FUNCTION_BLOCK FB_Gr01AutoAlarm
(*

The function block used to control alarms in manual mode.

Constructor: 		Patryk Panylo
Company:		E. Riexinger GmbH
Date:			28.04.2015
Version:			1.00

Date:			Revision:		Who:				Comment
dd.mm.yyyy		x.xx			Initials			comment

*)
VAR_INPUT
	(* Input variables / Eingang Variablen *)
	etMachineMode				:ET_MachineMode;			(* Machine mode *)
	etMachineState				:ET_MachineState;			(* Machine state *)
	bNoEStop					:BOOL;						(* Emergency stop *)
	bConfirmAlarm				:BOOL;						(* Confirm alarm *)
	dtDateTime 					:DATE_AND_TIME;			(* Actual date and time *)
	nFatalErrorMaxIdx				:INT;						(* Maximal index of  using alarms *)
	nErrorMaxIdx					:INT;						(* Maximal index of  using alarms *)
	nWarningMaxIdx				:INT;						(* Maximal index of  using alarms *)
	nMessageMaxIdx				:INT;						(* Maximal index of  using alarms *)
	nHintMaxIdx					:INT;						(* Maximal index of  using alarms *)
	stAlarmIn						:ST_AlarmIn;					(* Alarm input *)
END_VAR
VAR_OUTPUT
	(* Output variables / Ausgang Variablen *)
	stAlarmOut					:ST_AlarmOut;				(* Alarm input *)
END_VAR
VAR_IN_OUT
	(* Input Output variables / Ausgang Variablen *)
	bMoveInterrupted				:BOOL;						(* Move interrupted *)
	bHomeCompleted				:BOOL;						(* Home completed *)
END_VAR
VAR
	(* Enummerations *)

	(* Variables *)

	(* References *)

	(* Interfaces *)

	(* Instances *)
	fbAlarm						:FB_Alarm;
END_VAR


(* Collection of alarms *)
fbAlarm(
	bEnable := TRUE,
	bNoEStop := bNoEStop,
	bReset := bConfirmAlarm,
	dtDateTime := dtDateTime,
	nFatalErrorMaxIdx := nFatalErrorMaxIdx,
	nErrorMaxIdx := nErrorMaxIdx,
	nWarningMaxIdx := nWarningMaxIdx,
	nMessageMaxIdx := nMessageMaxIdx,
	nHintMaxIdx := nHintMaxIdx,
    	stAlarmIn := stAlarmIn,
    	stAlarmOut => stAlarmOut
);

IF stAlarmOut.bFatalError
    OR stAlarmOut.bError
THEN
	(*bMoveInterrupted := FALSE;*)
	bHomeCompleted := FALSE;
END_IF;

END_FUNCTION_BLOCK

(* stored: Version 1.1.0.1, ProductVersion 3.1.4024.15
   POU FB_Gr01AutoAlarm: Id {ff0c5e80-8dd8-4a8f-bdd6-61545f4a1244}, SpecialFunc None *)
